// TIA Portal project "Prova 1" (V17)

(* hardware
DEVICE "S7-1200 station_1"  S7-1200 Station
   slot 0: "Rack_0"  S7-1200 Rack  Rack  V1.0
   slot 1: "PLC_1"  CPU 1214C DC/DC/DC  6ES7 214-1AG31-0XB0  V3.0
*)

// ===== PLC "PLC_1"  CPU 1214C DC/DC/DC =====

VAR_GLOBAL   // PLC tag table "Default tag table"
   "Sensor_Indutivo_Leste (Home)" AT %I0.2 : Bool;
   "Sensor_Indutivo_Oeste" AT %I0.3 : Bool;
   "Sensor_Optico" AT %I0.4 : Bool;
   "Entrada_Encoder_A" AT %I0.0 : Bool;
   "Entrada_Encoder_B" AT %I0.1 : Bool;
   "Voltas" AT %ID1000 : DWord;
   "PUL" AT %Q0.0 : Bool;
   "DIR" AT %Q0.1 : Bool;
   "EN" AT %Q0.2 : Bool;
   "enable" AT %I0.5 : Bool;
   "saida" AT %Q0.3 : Bool;
   "Mover_Direita" AT %M10.0 : Bool;
   "Mover_Esquerda" AT %M10.1 : Bool;
   "Memória_Home" AT %M10.2 : Bool;
   "M_Subida" AT %M10.3 : Bool;
   "M_Subida2" AT %M10.4 : Bool;
   "M_Subida3" AT %M10.5 : Bool;
   "M_Subida4" AT %M10.6 : Bool;
   "Teste" AT %I0.6 : Bool;
   "Velovidade" AT %Q0.5 : Bool;
   "Gira/Para" AT %Q0.4 : Bool;
   "M_Subida5" AT %M10.7 : Bool;
   "Trepidar" AT %M11.0 : Bool;
   "System_Byte" AT %MB1 : Byte;
   "FirstScan" AT %M1.0 : Bool;
   "DiagStatusUpdate" AT %M1.1 : Bool;
   "AlwaysTRUE" AT %M1.2 : Bool;
   "AlwaysFALSE" AT %M1.3 : Bool;
   "Clock_Byte" AT %MB0 : Byte;
   "Clock_10Hz" AT %M0.0 : Bool;
   "Clock_5Hz" AT %M0.1 : Bool;
   "Clock_2.5Hz" AT %M0.2 : Bool;
   "Clock_2Hz" AT %M0.3 : Bool;
   "Clock_1.25Hz" AT %M0.4 : Bool;
   "Clock_1Hz" AT %M0.5 : Bool;
   "Clock_0.625Hz" AT %M0.6 : Bool;
   "Clock_0.5Hz" AT %M0.7 : Bool;
   "M_Subida6" AT %M11.1 : Bool;
   "M_Subida7" AT %M11.2 : Bool;
   "M_Subida8" AT %M11.3 : Bool;
   "Lavagem" AT %M11.4 : Bool;
   "Manutencao" AT %M11.5 : Bool;
   "Reparado" AT %I0.7 : Bool;
   "M_subida9" AT %M11.6 : Bool;
   "Reset voltas" AT %M11.7 : Bool;
   "M_subida10" AT %M12.0 : Bool;
END_VAR

DATA_BLOCK "Agendamento do Sol_DB"   // DB3
{ S7_Optimized_Access := 'TRUE' }
VERSION : 0.1
// stored: InstanceOfName Agendamento do Sol
"Agendamento do Sol"
BEGIN
END_DATA_BLOCK

DATA_BLOCK "Encoder"   // DB12
{ S7_Optimized_Access := 'TRUE' }
VERSION : 0.1
   VAR RETAIN
      Contagem_Valor : DInt;
   END_VAR
   VAR
      Referencia_Valor : DInt := 900;
      DIR : Bool;
      "Valor_(T-1)" : DInt;
   END_VAR
   VAR RETAIN
      "valor(T)" : DInt;
   END_VAR
   VAR
      Delta : DInt;
   END_VAR
BEGIN
END_DATA_BLOCK

DATA_BLOCK "Lavagem_Inversor_DB_1"   // DB15
{ S7_Optimized_Access := 'TRUE' }
VERSION : 0.1
// stored: InstanceOfName Lavagem_Inversor
"Lavagem_Inversor"
BEGIN
END_DATA_BLOCK

DATA_BLOCK "Controle Motor de Passo_DB_1"   // DB18
{ S7_Optimized_Access := 'TRUE' }
VERSION : 0.1
// stored: InstanceOfName Controle Motor de Passo
"Controle Motor de Passo"
BEGIN
END_DATA_BLOCK

// folder: System blocks/Program resources

DATA_BLOCK "IEC_Timer_0_DB"   // DB10
{ S7_Optimized_Access := 'TRUE' }
AUTHOR : Simatic
FAMILY : IEC
NAME : IEC_TMR
VERSION : 1.0
// stored: InstanceOfName IEC_TIMER
"IEC_TIMER"
BEGIN
END_DATA_BLOCK

DATA_BLOCK "IEC_Timer_0_DB_1"   // DB11
{ S7_Optimized_Access := 'TRUE' }
AUTHOR : Simatic
FAMILY : IEC
NAME : IEC_TMR
VERSION : 1.0
// stored: InstanceOfName IEC_TIMER
"IEC_TIMER"
BEGIN
END_DATA_BLOCK

// folder: (top level)

DATA_BLOCK "Axis_1"   // DB1, Motion_DB
{ S7_Optimized_Access := 'TRUE' }
AUTHOR : SIMATIC
FAMILY : BasicMC
NAME : TO_PTO
VERSION : 3.0
// stored: InstanceOfName TO_Axis_PTO
"TO_Axis_PTO"
BEGIN
   // Axis.LengthUnit.LastDistance = 1005
   // Axis.HomingReferencePointSwitch_AddressCU = %I0.2
   // Axis.LengthUnitNormalized.Distance = 1005
   // Axis.EnableOutput_AddressCU = %Q0.2
   // Axis.DirectionHwcnAddressCU = Q0.1
   // Axis.PulseHwcnAddressCU = Q0.0
   // Pulse.MinDeltaDeltaFrequencyCU = 0.004
   // Pulse.MaxDeltaDeltaFrequencyCU = 1.0E+10
   // Pulse.MinDeltaFrequencyCU = 0.005
   // Pulse.MaxDeltaFrequencyCU = 9.5E+9
   // Pulse.MinFrequencyCU = 1.0
   // Pulse.MaxFrequencyCU = 100000.0
   // Pulse.OutputSourceCU = 16#0000_0000
   // Axis.SelectPTO = 0
END_DATA_BLOCK

FUNCTION_BLOCK "Agendamento do Sol"   // FB1, LAD
{ S7_Optimized_Access := 'TRUE' }
VERSION : 0.1
   VAR_INPUT
      "Entrada Teste" : Bool;
   END_VAR
   VAR
      Tempo : DTL;
      Verifica : Int;
   END_VAR
BEGIN

REGION Network 1: Ler o Tempo_Atual
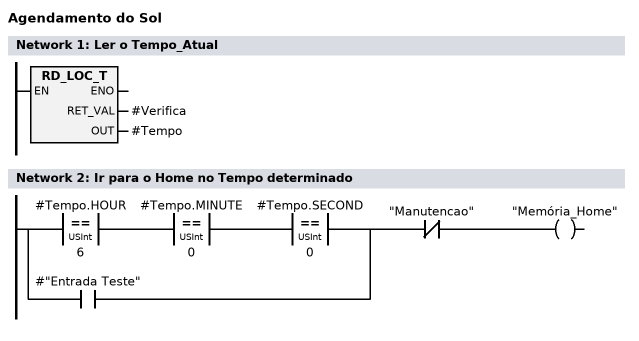
   #Verifica := RD_LOC_T(OUT => #Tempo);
END_REGION

REGION Network 2: Ir para o Home no Tempo determinado
   RUNG wire#powerrail
      { S7_Templates := "SrcType := USInt" } EQ_Contact(in1 := #Tempo.HOUR, in2 := 6)
      { S7_Templates := "SrcType := USInt" } EQ_Contact(in1 := #Tempo.MINUTE, in2 := 0)
      { S7_Templates := "SrcType := USInt" } EQ_Contact(in1 := #Tempo.SECOND, in2 := 0)
      wire#w1
      I_Contact( "Manutencao" )
      Coil( "Memória_Home" )
   END_RUNG
   RUNG wire#powerrail
      Contact( #"Entrada Teste" )
   END_RUNG wire#w1
   // the same network as SCL:
   "Memória_Home" := (((#Tempo.HOUR = 6) AND (#Tempo.MINUTE = 0) AND (#Tempo.SECOND = 0)) OR #"Entrada Teste") AND NOT "Manutencao";
END_REGION
END_FUNCTION_BLOCK

FUNCTION_BLOCK "Lavagem_Inversor"   // FB2, LAD
{ S7_Optimized_Access := 'TRUE' }
VERSION : 0.1
   VAR_INPUT
      Reparo : Bool;
   END_VAR
   VAR_TEMP   // added for the SCL form of the ladder/FBD networks
      _w1 : Bool;
   END_VAR
BEGIN

REGION Network 1: Começar Processo de Lavagem
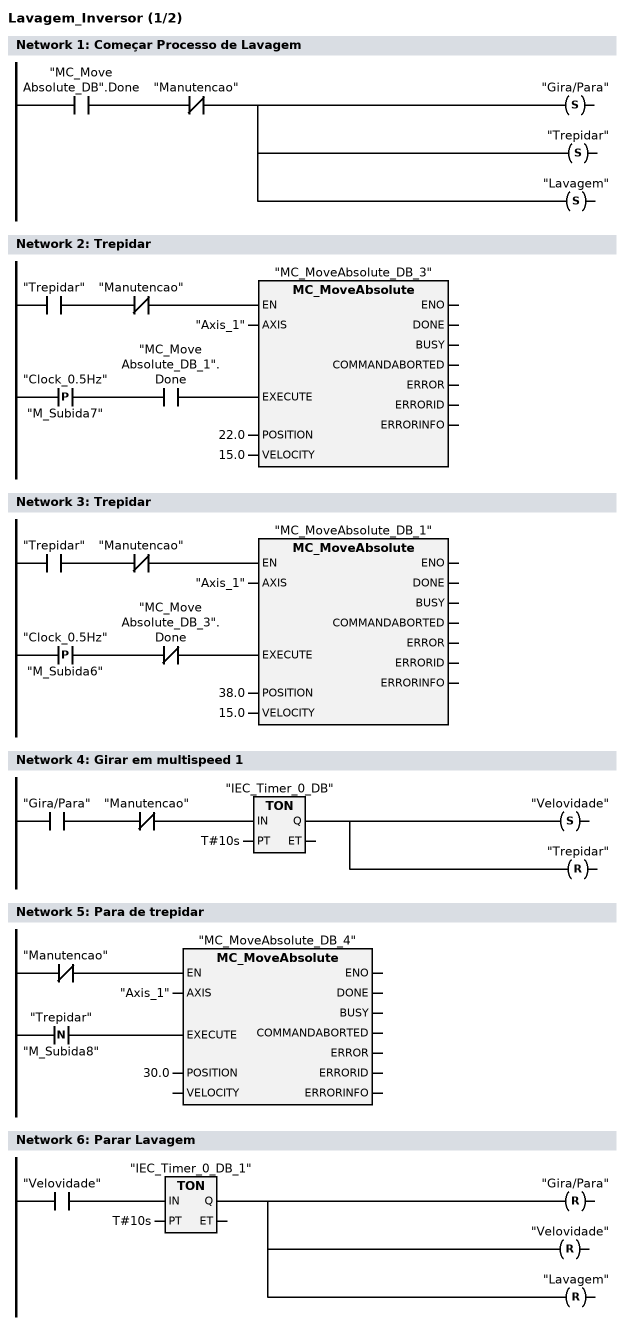
   RUNG wire#powerrail
      Contact( "MC_MoveAbsolute_DB".Done )
      I_Contact( "Manutencao" )
      wire#w1
      S_Coil( "Gira/Para" )
   END_RUNG
   RUNG wire#w1
      S_Coil( "Trepidar" )
   END_RUNG
   RUNG wire#w1
      S_Coil( "Lavagem" )
   END_RUNG
   // the same network as SCL:
   IF "MC_MoveAbsolute_DB".Done AND NOT "Manutencao" THEN
       "Gira/Para" := TRUE;
       "Trepidar" := TRUE;
       "Lavagem" := TRUE;
   END_IF;
END_REGION

REGION Network 2: Trepidar
   #_w1 := "Clock_0.5Hz" AND NOT "M_Subida7";   // rising edge of "Clock_0.5Hz"
   "M_Subida7" := "Clock_0.5Hz";
   IF "Trepidar" AND NOT "Manutencao" THEN
       "MC_MoveAbsolute_DB_3"(Axis := "Axis_1",   // MC_MoveAbsolute
                              Execute := #_w1 AND "MC_MoveAbsolute_DB_1".Done,
                              Position := 22.0,
                              Velocity := 15.0);
   END_IF;
END_REGION

REGION Network 3: Trepidar
   #_w1 := "Clock_0.5Hz" AND NOT "M_Subida6";   // rising edge of "Clock_0.5Hz"
   "M_Subida6" := "Clock_0.5Hz";
   IF "Trepidar" AND NOT "Manutencao" THEN
       "MC_MoveAbsolute_DB_1"(Axis := "Axis_1",   // MC_MoveAbsolute
                              Execute := #_w1 AND NOT "MC_MoveAbsolute_DB_3".Done,
                              Position := 38.0,
                              Velocity := 15.0);
   END_IF;
END_REGION

REGION Network 4: Girar em multispeed 1
   "IEC_Timer_0_DB".TON(IN := "Gira/Para" AND NOT "Manutencao", PT := T#10s);
   IF "IEC_Timer_0_DB".Q THEN
       "Velovidade" := TRUE;
       "Trepidar" := FALSE;
   END_IF;
END_REGION

REGION Network 5: Para de trepidar
   #_w1 := NOT "Trepidar" AND "M_Subida8";   // falling edge of "Trepidar"
   "M_Subida8" := "Trepidar";
   IF NOT "Manutencao" THEN
       "MC_MoveAbsolute_DB_4"(Axis := "Axis_1", Execute := #_w1, Position := 30.0);   // MC_MoveAbsolute
   END_IF;
END_REGION

REGION Network 6: Parar Lavagem
   "IEC_Timer_0_DB_1".TON(IN := "Velovidade", PT := T#10s);
   IF "IEC_Timer_0_DB_1".Q THEN
       "Gira/Para" := FALSE;
       "Velovidade" := FALSE;
       "Lavagem" := FALSE;
   END_IF;
END_REGION

REGION Network 7: Voltar para posicao alvorada
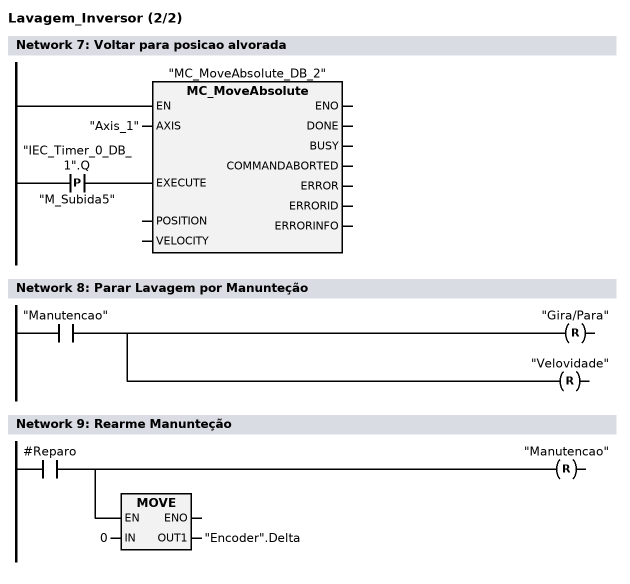
   #_w1 := "IEC_Timer_0_DB_1".Q AND NOT "M_Subida5";   // rising edge of "IEC_Timer_0_DB_1".Q
   "M_Subida5" := "IEC_Timer_0_DB_1".Q;
   "MC_MoveAbsolute_DB_2"(Axis := "Axis_1", Execute := #_w1);   // MC_MoveAbsolute
END_REGION

REGION Network 8: Parar Lavagem por Manunteção
   RUNG wire#powerrail
      Contact( "Manutencao" )
      wire#w1
      R_Coil( "Gira/Para" )
   END_RUNG
   RUNG wire#w1
      R_Coil( "Velovidade" )
   END_RUNG
   // the same network as SCL:
   IF "Manutencao" THEN
       "Gira/Para" := FALSE;
       "Velovidade" := FALSE;
   END_IF;
END_REGION

REGION Network 9: Rearme Manunteção
   RUNG wire#powerrail
      Contact( #Reparo )
      wire#w1
      R_Coil( "Manutencao" )
   END_RUNG
   RUNG wire#w1
      { S7_GenerateENO := "TRUE" } Move(in := 0, out1 => "Encoder".Delta)
   END_RUNG
   // the same network as SCL:
   IF #Reparo THEN
       "Manutencao" := FALSE;
       "Encoder".Delta := 0;
   END_IF;
END_REGION
END_FUNCTION_BLOCK

FUNCTION_BLOCK "Controle Motor de Passo"   // FB3, LAD
{ S7_Optimized_Access := 'TRUE' }
VERSION : 0.1
   VAR_INPUT
      "Entrada do Sensor" : Bool;
   END_VAR
   VAR_TEMP   // added for the SCL form of the ladder/FBD networks
      _w1 : Bool;
   END_VAR
BEGIN

REGION Network 1: Ativar Motor
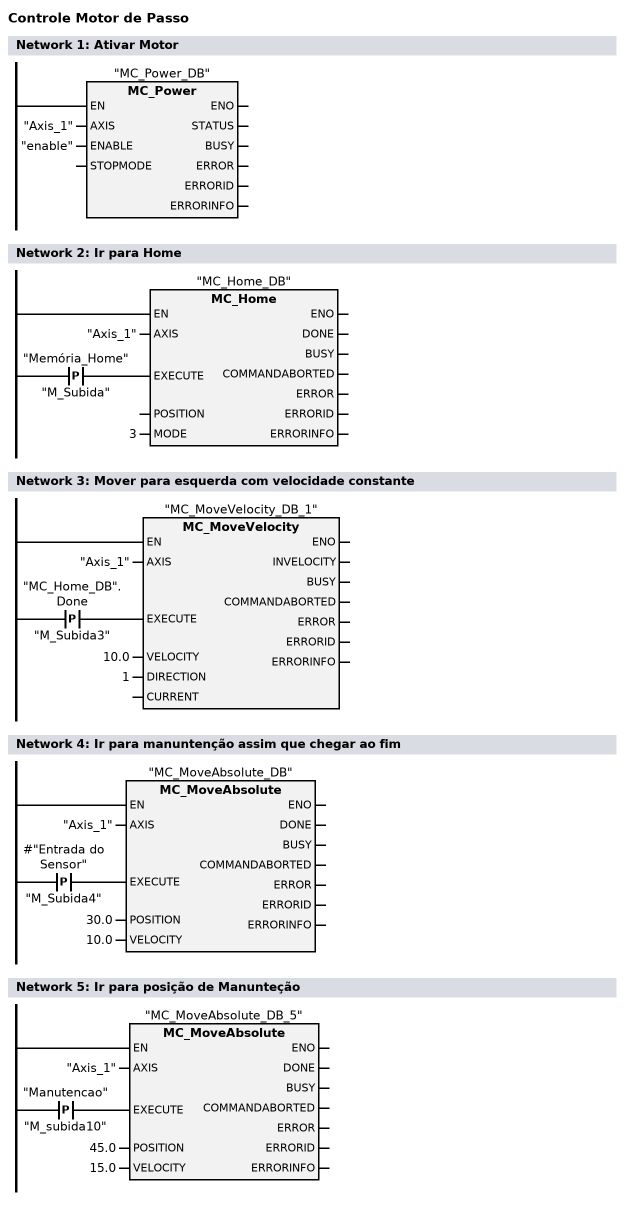
   "MC_Power_DB"(Axis := "Axis_1", Enable := "enable");   // MC_Power
END_REGION

REGION Network 2: Ir para Home
   #_w1 := "Memória_Home" AND NOT "M_Subida";   // rising edge of "Memória_Home"
   "M_Subida" := "Memória_Home";
   "MC_Home_DB"(Axis := "Axis_1", Execute := #_w1, Mode := 3);   // MC_Home
END_REGION

REGION Network 3: Mover para esquerda com velocidade constante
   #_w1 := "MC_Home_DB".Done AND NOT "M_Subida3";   // rising edge of "MC_Home_DB".Done
   "M_Subida3" := "MC_Home_DB".Done;
   "MC_MoveVelocity_DB_1"(Axis := "Axis_1", Execute := #_w1, Velocity := 10.0, Direction := 1);   // MC_MoveVelocity
END_REGION

REGION Network 4: Ir para manuntenção assim que chegar ao fim
   #_w1 := #"Entrada do Sensor" AND NOT "M_Subida4";   // rising edge of #"Entrada do Sensor"
   "M_Subida4" := #"Entrada do Sensor";
   "MC_MoveAbsolute_DB"(Axis := "Axis_1", Execute := #_w1, Position := 30.0, Velocity := 10.0);   // MC_MoveAbsolute
END_REGION

REGION Network 5: Ir para posição de Manunteção
   #_w1 := "Manutencao" AND NOT "M_subida10";   // rising edge of "Manutencao"
   "M_subida10" := "Manutencao";
   "MC_MoveAbsolute_DB_5"(Axis := "Axis_1", Execute := #_w1, Position := 45.0, Velocity := 15.0);   // MC_MoveAbsolute
END_REGION
END_FUNCTION_BLOCK

FUNCTION "Encoder Fc" : Void   // FC1, LAD
{ S7_Optimized_Access := 'TRUE' }
VERSION : 0.1
   VAR_TEMP   // added for the SCL form of the ladder/FBD networks
      _w1 : Bool;
   END_VAR
BEGIN

REGION Network 1
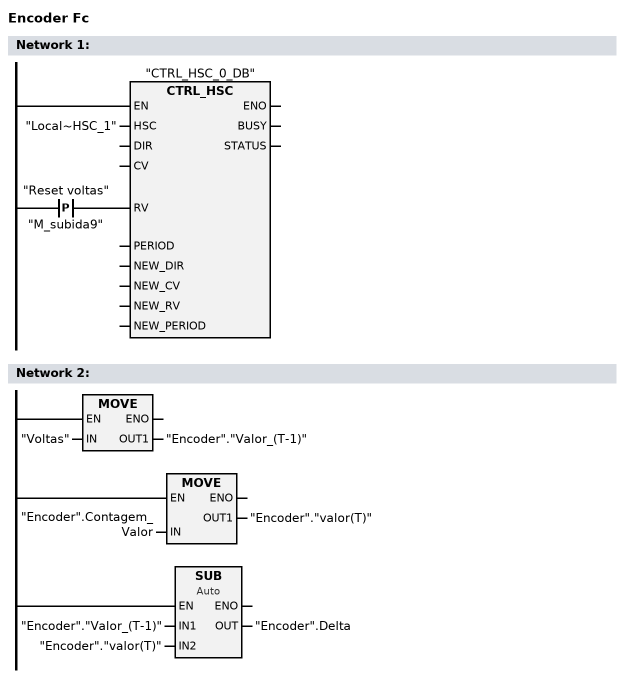
   #_w1 := "Reset voltas" AND NOT "M_subida9";   // rising edge of "Reset voltas"
   "M_subida9" := "Reset voltas";
   "CTRL_HSC_0_DB"(HSC := "Local~HSC_1", RV := #_w1);   // CTRL_HSC
END_REGION

REGION Network 2
   RUNG wire#powerrail
      { S7_GenerateENO := "TRUE" } Move(in := "Voltas", out1 => "Encoder"."Valor_(T-1)")
   END_RUNG
   RUNG wire#powerrail
      { S7_GenerateENO := "TRUE" } Move(in := "Encoder".Contagem_Valor, out1 => "Encoder"."valor(T)")
   END_RUNG
   RUNG wire#powerrail
      { S7_GenerateENO := "TRUE" } Sub(in1 := "Encoder"."Valor_(T-1)", in2 := "Encoder"."valor(T)", out => "Encoder".Delta)
   END_RUNG
   // the same network as SCL:
   "Encoder"."Valor_(T-1)" := "Voltas";
   "Encoder"."valor(T)" := "Encoder".Contagem_Valor;
   "Encoder".Delta := "Encoder"."Valor_(T-1)" - "Encoder"."valor(T)";
END_REGION
END_FUNCTION

ORGANIZATION_BLOCK "Main"   // OB1, LAD, ProgramCycle
TITLE = "Main Program Sweep (Cycle)"
{ S7_Optimized_Access := 'TRUE' }
VERSION : 0.1
BEGIN

REGION Network 1: Ler o Tempo_Atual
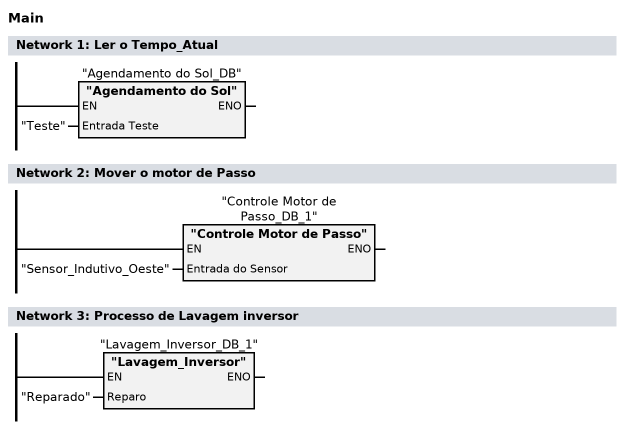
   RUNG wire#powerrail
      "Agendamento do Sol_DB"("Entrada Teste" := "Teste")
   END_RUNG
   // the same network as SCL:
   "Agendamento do Sol_DB"("Entrada Teste" := "Teste");   // "Agendamento do Sol"
END_REGION

REGION Network 2: Mover o motor de Passo
   RUNG wire#powerrail
      "Controle Motor de Passo_DB_1"("Entrada do Sensor" := "Sensor_Indutivo_Oeste")
   END_RUNG
   // the same network as SCL:
   "Controle Motor de Passo_DB_1"("Entrada do Sensor" := "Sensor_Indutivo_Oeste");   // "Controle Motor de Passo"
END_REGION

REGION Network 3: Processo de Lavagem inversor
   RUNG wire#powerrail
      "Lavagem_Inversor_DB_1"(Reparo := "Reparado")
   END_RUNG
   // the same network as SCL:
   "Lavagem_Inversor_DB_1"(Reparo := "Reparado");   // "Lavagem_Inversor"
END_REGION
END_ORGANIZATION_BLOCK

ORGANIZATION_BLOCK "Interrupção encoder"   // OB40, LAD, HWProcessInterrupt
{ S7_Optimized_Access := 'TRUE' }
VERSION : 0.1
   VAR_TEMP   // added for the SCL form of the ladder/FBD networks
      _w1 : Bool;
   END_VAR
BEGIN

REGION Network 1: Intertravamento
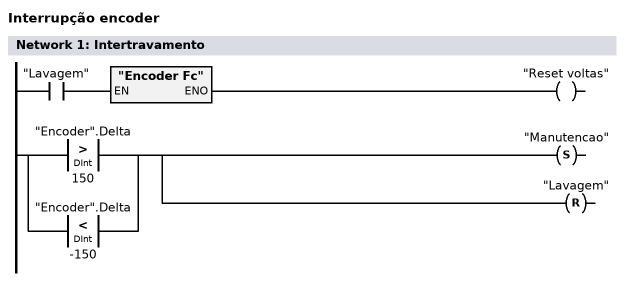
   RUNG wire#powerrail
      Contact( "Lavagem" )
      "Encoder Fc"()
      Coil( "Reset voltas" )
   END_RUNG
   RUNG wire#powerrail
      { S7_Templates := "SrcType := DInt" } GT_Contact(in1 := "Encoder".Delta, in2 := 150)
      wire#w1
      S_Coil( "Manutencao" )
   END_RUNG
   RUNG wire#powerrail
      { S7_Templates := "SrcType := DInt" } LT_Contact(in1 := "Encoder".Delta, in2 := -150)
   END_RUNG wire#w1
   RUNG wire#w1
      R_Coil( "Lavagem" )
   END_RUNG
   // the same network as SCL:
   "Encoder Fc"(EN := "Lavagem", ENO => #_w1);
   "Reset voltas" := #_w1;
   IF ("Encoder".Delta > 150) OR ("Encoder".Delta < (-150)) THEN
       "Manutencao" := TRUE;
       "Lavagem" := FALSE;
   END_IF;
END_REGION
END_ORGANIZATION_BLOCK